// TIA Portal V21 export
// export: Created 2026-10-14T03:11:20.9082904Z, ExportSetting WithDefaults, DisplayName Totally Integrated Automation Portal, DisplayVersion V21, DisplayName STEP 7 Professional, DisplayVersion V21, DisplayName STEP 7 Safety, DisplayVersion V21, DisplayName Tech WebApplication, DisplayVersion V21, DisplayName WinCC Basic/Comfort/Advanced, DisplayVersion V21, DisplayName WinCC Unified, DisplayVersion V21
TagTable "LCCA_PvSim_PID_C"
  LLCCA_PvSim_PID_C_DB_enable : Bool  (HMI_Connection_1, 1 s)
  LLCCA_PvSim_PID_C_DB_input : Real  (HMI_Connection_1, 100 ms)
  LLCCA_PvSim_PID_C_DB_out : Real  (HMI_Connection_1, 100 ms)
  LLCCA_PvSim_PID_C_DB_addComp : Real  (HMI_Connection_1, 100 ms)
  LLCCA_PvSim_PID_C_DB_subComp : Real  (HMI_Connection_1, 100 ms)
  LLCCA_PvSim_PID_C_DB_reset : Bool  (HMI_Connection_1, 1 s)
  LLCCA_PvSim_PID_C_DB_ioAddFactor : Real  (HMI_Connection_1, 1 s)
  LLCCA_PvSim_PID_C_DB_ioAddTimeLag : USInt  (HMI_Connection_1, 1 s)
  LLCCA_PvSim_PID_C_DB_ioAddFilter : Real  (HMI_Connection_1, 1 s)
  LLCCA_PvSim_PID_C_DB_ioSubFactor : Real  (HMI_Connection_1, 1 s)
  LLCCA_PvSim_PID_C_DB_ioSubStartValue : Real  (HMI_Connection_1, 1 s)
  LLCCA_PvSim_PID_C_DB_ioNoiceFactor : Real  (HMI_Connection_1, 1 s)
  LLCCA_PvSim_PID_C_DB_ioSubConstant : Real  (HMI_Connection_1, 1 s)
  LLCCA_PvSim_PID_C_DB_ioSubType : USInt  (HMI_Connection_1, 1 s)
  LLCCA_PvSim_PID_C_DB_ioSubTimeLag : USInt  (HMI_Connection_1, 1 s)
  LLCCA_PvSim_PID_C_DB_ioSubFilter : Real  (HMI_Connection_1, 1 s)
